// TIA Portal V19 export
TYPE "UDT_TachoDT_I"
   STRUCT
      ZSO_112B : Bool;
      ZSO_112A : Bool;
      ZSO_105 : Bool;
      ZSO_103 : Bool;
      ZSO_109 : Bool;
      ZSO_104 : Bool;
      ZSO_108 : Bool;
      YI_101 : Bool;   // Agitador en marcha
      YT_101 : Bool;   // Disparo del agitador
      ZSO_102 : Bool;
      ZSO_113 : Bool;
      YI_102 : Bool;   // Bomba de vacÃ­o en marcha Entradas analÃ³gicas: RAW 0..27648
      LT_112_RAW : Int;
      PT_110_RAW : Int;
      PT_113_RAW : Int;
      TT_114_RAW : Int;
      TT_115_RAW : Int;
      AT_112_RAW : Int;
      LT_116_RAW : Int;
      AT_112X_RAW : Int;
   END_STRUCT;
END_TYPE
